PROGRAM MAIN
VAR
    iCount : INT;
    bLight : BOOL;
    bSwitch : BOOL;
END_VAR

iCount := iCount + 1;

// reset logic
IF iCount > 100 THEN
    iCount := 0;
END_IF

// new Light/Switch logic
IF iCount > 50 THEN
    bLight := bSwitch;
ELSE
    bLight := FALSE;
END_IF

END_PROGRAM

(* stored: Version 1.1.0.1
   POU MAIN: Id {a48d85b8-1883-40f5-b698-0e9758ed2b9e}, SpecialFunc None *)
